// TIA Portal V21 export
// export: Created 2026-11-11T00:47:47.1876166Z, ExportSetting WithDefaults, DisplayName Totally Integrated Automation Portal, DisplayVersion V21 Update 3, DisplayName STEP 7 Professional, DisplayVersion V21 Update 3, DisplayName STEP 7 Safety, DisplayVersion V21, DisplayName Tech WebApplication, DisplayVersion V21, DisplayName WinCC Basic/Comfort/Advanced, DisplayVersion V21 Update 3, DisplayName WinCC Unified, DisplayVersion V21 Update 3
FUNCTION_BLOCK "FB_Fbd_sc004"   // FB183, FBD
{ S7_Optimized_Access := 'TRUE' }
VERSION : 0.1
// stored: AutoNumber true, IsIECCheckEnabled false, IsRetainMemResEnabled false, MemoryReserve 100, SetENOAutomatically false, UDAEnableTagReadback false
   VAR_INPUT
      v_en_r : Bool;
      v_id : CONN_PRG;
      v_r_id : CONN_R_ID;
   END_VAR
   VAR_OUTPUT
      v_ndr : Bool;
      v_error : Bool;
      v_status : Word;
   END_VAR
   VAR_IN_OUT
      v_rd_1 : Variant;
      v_rd_2 : Variant;
      v_rd_3 : Variant;
      v_rd_4 : Variant;
   END_VAR
   VAR
      inst { S7_SetPoint := 'True'} : URCV;
   END_VAR
BEGIN

REGION Network 1: URCV - Receive data uncoordinated
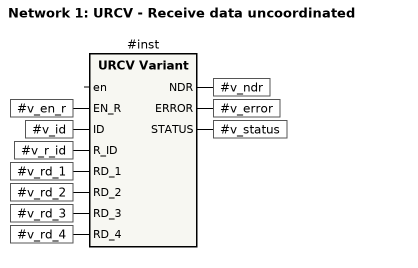
   #inst(EN_R := #v_en_r,   // URCV
         ID := #v_id,
         R_ID := #v_r_id,
         RD_1 := #v_rd_1,
         RD_2 := #v_rd_2,
         RD_3 := #v_rd_3,
         RD_4 := #v_rd_4,
         NDR => #v_ndr,
         ERROR => #v_error,
         STATUS => #v_status);
END_REGION
END_FUNCTION_BLOCK
